Fanuc KAREL source: kt00366.KL

-- PROVISIONAL review KL for V1013-1; original PC SHA256 e0bf836e2c0548b04439eb1eaca726f311c1ffc72eee963d07fda3c961d0f4ae
-- Incomplete behavior may be omitted. Consult companion uncertainty JSON. Do not deploy.
PROGRAM KT00366
%NOLOCKGROUP
VAR
  I1 : INTEGER
  R2 : REAL
  OUT : BOOLEAN
BEGIN
  -- UNRESOLVED_PC offsets 5-16; opcodes 2E,23
  -- UNRESOLVED_PC offsets 21-32; opcodes 2E,23
  -- UNRESOLVED_PC offsets 37-59; opcodes 21,21,29,64,29,70,23
  -- UNRESOLVED_PC offsets 64-68; opcodes 7F
END KT00366
